// TIA Portal V19 export
DATA_BLOCK "iRC_Pick_R2"   // DB7
// stored: InstanceOfName RC_Pick, InstanceOfType FB
"RC_Pick"
   // VAR_INPUT
   //    Execute : Bool;
   // END_VAR
   // VAR_OUTPUT
   //    Busy : Bool;
   //    Done : Bool;
   //    Error : Bool;
   //    ErrorId : Int;
   // END_VAR
   // VAR_IN_OUT
   //    Robot : "ST_ROBOT";
   // END_VAR
   // VAR
   //    iStage : Int;
   //    iRC_CallProgramm : "RC_CallProgram";
   //    xGo { S7_SetPoint := 'True'} : Bool;
   // END_VAR
BEGIN
END_DATA_BLOCK
